Universal Robots PolyScope program: ApproachMove.urp

Program ApproachMove (createdIn=3.0.0 lastSavedIn=3.0.0 directory=/programs installation=default)
Robot Program (runOnlyOnce=true motionType=MoveJ speed=1.047198 acceleration=1.396263 useActiveTCP=false)
  'Program generated by VerticalBot Studio for UR10 on 25/10/2026 12:00:00'
  'Using nominal kinematics.'
  'Using Ref. Frame 2: p[-0.800000, 0.500000, 0.100000, 0.000000, 0.000000, 3.141593]'
  'Using TCP Paint gun: p[0.050000, 0.000000, 0.450000, 0.000000, 0.523599, 0.000000]'
  Script: set_tcp(p[0.050000, 0.000000, 0.450000, 0.000000, 0.523599, 0.000000])
  Script: movej([-2.652656, -1.365240, -1.512183, -1.127521, 1.275171, 1.920421],1.20000,0.75000,0,0.0000)
  MoveJ speed 42.97 deg/s, acceleration 68.75 deg/s^2 (useActiveTCP=true)
    Waypoint Waypoint_1: TCP in base x=-866.761 y=-115.117 z=513.712 mm, rx=3.1014 ry=0.052 rz=-0.3627 rad; joints [-151.986, -78.222, -86.642, -64.602, 73.062, 110.032] deg; flange x=-594.55 y=-100.237 z=875.208 mm, rx=2.8946 ry=0.0426 rz=-1.1501 rad
  Script: movej([-3.642345, -1.680989, -1.433833, -1.128762, 1.813205, 1.128191],1.20000,0.75000,0,0.0000)
  MoveJ speed 42.97 deg/s, acceleration 68.75 deg/s^2 (useActiveTCP=true)
    Waypoint Waypoint_2: TCP in base x=-800 y=500 z=300 mm, rx=3.1416 ry=0 rz=0 rad; joints [-208.691, -96.314, -82.153, -64.673, 103.889, 64.641] deg; flange x=-618.301 y=500 z=714.711 mm, rx=3.0345 ry=0 rz=-0.8131 rad
